// TIA Portal V20 export
TYPE "WT3_HoldingRegister_UDT"
   STRUCT
      Index : Array[1..32767] of Word;   // 32767 Words (Max 65'532‬ Bytes)
   END_STRUCT;
END_TYPE
